{attribute 'linkalways'} 
{attribute 'no_explicit_call' := 'This FB is a CLASS and must be accessed using methods or properties'}
{attribute 'enable_dynamic_creation'}
FUNCTION_BLOCK _Array0to2OfLREAL EXTENDS ArrayDatatypeBase_1D
VAR CONSTANT
	lBound : DINT := 0;
	uBound : DINT := 2;
END_VAR
VAR
	localData : ARRAY [lBound..uBound] OF LREAL;
	activeData : REFERENCE TO ARRAY [lBound..uBound] OF LREAL REF= localData;
	elements : ARRAY [lBound..uBound] OF _LREAL(0.0);
	baseType : _LREAL(0.0);
END_VAR

PROPERTY PUBLIC Address : PVOID
GET
Address := ADR(activeData);
END_GET
END_PROPERTY

PROPERTY PUBLIC BaseDatatype : I_Datatype
GET
BaseDatatype := baseType;
END_GET
END_PROPERTY

METHOD PUBLIC ClearReference
VAR_INPUT
END_VAR
activeData REF= localData;
SetElementReference();
END_METHOD

METHOD PUBLIC Clone : I_Datatype
VAR
    pClone : POINTER TO _Array0to2OfLREAL;
END_VAR
pClone := __NEW(_Array0to2OfLREAL());
pClone^.Value := Value;
Clone := pClone^;
END_METHOD

METHOD FB_init : BOOL
VAR_INPUT
	bInitRetains : BOOL; // if TRUE, the retain variables are initialized (warm start / cold start)
	bInCopyCode : BOOL;  // if TRUE, the instance afterwards gets moved into the copy code (online change)
END_VAR
SetElementReference();
END_METHOD

METHOD PUBLIC MakeReferenceTo
VAR_INPUT
	ReferenceTarget : REFERENCE TO ARRAY [lBound..uBound] OF LREAL;
END_VAR
activeData REF= ReferenceTarget;
SetElementReference();
END_METHOD

METHOD PROTECTED OnSerializeArrayValues
VAR_INPUT
	Serializer : I_Serializer;
END_VAR
VAR
	i : DINT;
END_VAR
FOR i := lBound TO uBound DO
	elements[i].SerializeWith(Serializer);
END_FOR
END_METHOD

METHOD PROTECTED SetElementReference
VAR_INPUT
END_VAR
VAR
	i : DINT;
END_VAR
FOR i := lBound TO uBound DO
	elements[i].MakeReferenceTo(activeData[i]);
END_FOR
END_METHOD

PROPERTY PUBLIC Size : UDINT
GET
Size := SIZEOF(activeData);
END_GET
END_PROPERTY

METHOD PROTECTED TryDeserializeArrayValues : BOOL
VAR_INPUT
	Deserializer : I_Deserializer;
	Feedback : I_DeserializerFeedback;
END_VAR
VAR
	failed : BOOL;
	enumerator : I_DeserializerArrayForwardEnumerator;
	i : DINT;
END_VAR
enumerator := Deserializer.GetArrayEnumerator();
i := lBound;

WHILE enumerator.MoveNext() AND i <= uBound AND NOT failed DO
	
	IF NOT elements[i].TryDeserializeFrom(enumerator.Current, Feedback) THEN
		failed := TRUE;
		EXIT;
	END_IF
	i := i + 1;

END_WHILE
enumerator.Dispose();

TryDeserializeArrayValues := NOT failed;
END_METHOD

METHOD PUBLIC TryGetElementAsDatatypeByIndex : BOOL
VAR_INPUT
	Index : DINT;
	Destination : REFERENCE TO I_Datatype;
END_VAR
IF Index < lbound OR Index > ubound THEN
	RETURN;
END_IF

Destination := elements[Index];
TryGetElementAsDatatypeByIndex := TRUE;
END_METHOD

METHOD PUBLIC TryGetLowerBound : BOOL
VAR_INPUT
	Dimention : UDINT;
	Destination : REFERENCE TO DINT;
END_VAR
IF Dimention = 1 THEN
	Destination := lBound;
	TryGetLowerBound := TRUE;
END_IF
END_METHOD

METHOD PUBLIC TryGetUpperBound : BOOL
VAR_INPUT
	Dimention : UDINT;
	Destination : REFERENCE TO DINT;
END_VAR
IF Dimention = 1 THEN
	Destination := uBound;
	TryGetUpperBound := TRUE;
END_IF
END_METHOD

METHOD TryMakeReferenceTo : BOOL
VAR_INPUT
	Target : I_Datatype;
END_VAR
VAR
	pTargetData : POINTER TO ARRAY [lBound..uBound] OF LREAL;
END_VAR
IF NOT IsEquivalentTo(Target) THEN
	RETURN;
END_IF

pTargetData := Target.Address;
activeData REF= pTargetData^;
SetElementReference();
TryMakeReferenceTo := TRUE;
END_METHOD

PROPERTY PUBLIC Value : REFERENCE TO ARRAY [lBound..uBound] OF LREAL;
GET
Value ref= activeData;
END_GET
END_PROPERTY

END_FUNCTION_BLOCK

(* stored: Version 1.1.0.1, ProductVersion 3.1.4024.13
   POU _Array0to2OfLREAL: Id {9d380b32-3610-0bc4-2019-6c5e25a3aa16}, SpecialFunc None
   Folder Core: Id {9818e471-bbe5-0e2b-0f38-c1bcf2245d92}
   Folder Constructor: Id {6f413ee4-d95c-0694-011a-ebf1f51148b6}
   Folder Protected: Id {d9013ca9-3741-0110-30b5-46531f7b4912}
   Folder Customize: Id {f2870487-a827-004a-287a-ceb27a21e64b}
   Property Address: Id {029fb2f4-4806-0b23-2301-29260ed79269}
   Get Get: Id {a3fd2c39-8bfc-08ca-04f0-e14a046ad1ae}
   Property BaseDatatype: Id {b85615ec-e67d-06ca-0be2-c59bafe386ba}
   Get Get: Id {cf23c015-a348-0b71-24a8-fc0b60392738}
   Method ClearReference: Id {d239279b-1c64-075a-32d1-85c896634ac8}
   Method Clone: Id {8a98e5e4-6b48-0979-0473-baf08bcf9e97}
   Method FB_init: Id {09a5f170-8c25-0781-1ed6-705f3ee1ef1b}
   Method MakeReferenceTo: Id {12c17128-655e-001d-174a-a2b61e4307fc}
   Method OnSerializeArrayValues: Id {e7daf2aa-a188-04a6-2ff5-18daca3326c0}
   Method SetElementReference: Id {89c20fcc-1441-0f43-0561-754b181fcd6d}
   Property Size: Id {2893a7c8-253d-01dc-2ca3-dfefca16197d}
   Get Get: Id {96976844-e447-0754-1c59-ded97ee96d2b}
   Method TryDeserializeArrayValues: Id {a8556c52-9653-06b5-07b6-69a02f0be509}
   Method TryGetElementAsDatatypeByIndex: Id {095d4b68-d998-0ba7-0932-8519902c967b}
   Method TryGetLowerBound: Id {f1fce5e9-261a-023b-26c6-bdd3665e9bfd}
   Method TryGetUpperBound: Id {b4879b8e-228c-0631-2659-133872148b4e}
   Method TryMakeReferenceTo: Id {9405b493-b3cf-00bb-3c87-a780d9ce003c}
   Property Value: Id {fd14ec9b-ce94-0bf9-1948-24fcf47478f2}
   Get Get: Id {c1dccd54-0277-0a0d-1afe-ee7ee37a01c3} *)
